FUNCTION "Set_Bit_F"   // FC 7, author

VAR_INPUT
   Bit : UInt;
END_VAR

VAR_IN_OUT
   Var : Word;
END_VAR

   // RETURN : Void
BEGIN
    // Set the bit
    #Var := #Var OR SHL(IN := WORD#1, N := #Bit);

END_FUNCTION